Fanuc KAREL source: kb00009.KL

-- PROVISIONAL review KL for V770-1; original PC SHA256 af432d9f0f8a92a18ed3c9554103a8b60054e6e080667dd819d79fdd5eef083e
-- Incomplete behavior may be omitted. Consult companion uncertainty JSON. Do not deploy.
PROGRAM KB00009
%NOLOCKGROUP
VAR
  P1 : REAL
  P2 : REAL
  RESULT : REAL
BEGIN
  -- UNRESOLVED_PC offsets 5-16; opcodes 2E,23
  -- UNRESOLVED_PC offsets 21-32; opcodes 2E,23
  -- UNRESOLVED_PC offsets 37-58; opcodes 27,22,22,76,23
  -- UNRESOLVED_PC offsets 63-67; opcodes 7F
END KB00009
